Staubli VAL3: bind.pgx

public program bind()
  local string l_scbx
  local num l_i
  local string l_snum
  local string l_schk
begin
  //cbxlist
  userPageBind("action","cbxlist","options",sActionList,size(sActionList),"r")
  //cbx0
  //  for l_i = 0 to 5
  //    l_scbx="cbx"+toString("",l_i)
  //  userPageBind("action","cbx0","options",sIOList,49,"r")
  //  userPageBind("action","cbx1","options",sIOList,49,"r")
  //  userPageBind("action","cbx2","options",sIOList,49,"r")
  //  userPageBind("action","cbx3","options",sIOList,49,"r")
  //  userPageBind("action","cbx4","options",sIOList,49,"r")
  //  userPageBind("action","cbx5","options",sIOList,49,"r")
  //endFor
  //value
  userPageBind("action","cbxlist","value",sSelList,1,"rw")
  //
  for l_i = 0 to 5
    l_scbx="cbx"+toString("",l_i)
    userPageBind("action",l_scbx,"value",sSelIO[l_i],1,"rw")
    l_scbx="cbx"+toString("",10+l_i)
    userPageBind("action",l_scbx,"value",aEditItem.aActItem[l_i].sIOtype,1,"rw")
    l_scbx="cbx"+toString("",20+l_i)
    userPageBind("action",l_scbx,"value",aEditItem.aActItem[l_i].sValue,1,"rw")
  endFor
  //text
  userPageBind("action","txt1","value",aEditItem.sComment,1,"rw")
  //
  //num input
  for l_i = 0 to 5
    l_snum="nmb"+toString("",l_i)
    userPageBind("action",l_snum,"value",aEditItem.aActItem[l_i].nPulseValue,1,"rw")
  endFor

  //click
  userPageBindClick("action","btnback",bBack,true)
  userPageBindClick("action","btn1",bConfirm,true)
  //check
  for l_i = 0 to 5
    l_schk="chk"+toString("",l_i)
    userPageBind("action",l_schk,"checked",aEditItem.aActItem[l_i].bActive,1,"rw")
  endFor
end
